Fanuc KAREL source: kc00051.KL

-- PROVISIONAL review KL for V940-1; original PC SHA256 62e1cba9f6348f84c1fd032b7c012092202f5e2c8dda128fd048dab9e5a6f124
-- Incomplete behavior may be omitted. Consult companion uncertainty JSON. Do not deploy.
PROGRAM KC00051
%NOLOCKGROUP
BEGIN
  -- V9_ZERO_TABLE_METADATA_HINT layout=0002_ascii; no indexed target words; source/name/runtime held
  -- UNRESOLVED_PC offsets 5-29; opcodes 27,22,22,2A,22,31
  -- UNRESOLVED_PC offsets 34-38; opcodes 7F
END KC00051
